(* PLC project Palletizer_Cell4.project, CODESYS CODESYS V3.5 SP19 Patch 2 *)
(* stored: creationDateTime 2026-10-30T09:14:22.5521931, modificationDateTime 2026-10-30T09:13:58.1180274 *)

(* Palletizer cell state *)
{attribute 'strict'}
TYPE E_CellState : (Idle := 0, Homing := 1, Picking := 2, Placing := 3, Faulted := 99) INT;
END_TYPE

TYPE ST_Recipe : STRUCT
  sName : STRING(40);  (* Recipe name *)
  iLayers : INT;  (* Layers per pallet *)
  iBoxesPerLayer : INT;
  lrLayerHeight : LREAL;  (* mm *)
  ltSettle : LTIME;  (* Settle time after place *)
END_STRUCT;
END_TYPE

TYPE U_StatusWord : union;
END_TYPE

INTERFACE I_Station
END_INTERFACE

FUNCTION_BLOCK ABSTRACT FB_Station IMPLEMENTS I_Station
VAR_INPUT
	bEnable : BOOL;
END_VAR
VAR_OUTPUT
	bReady : BOOL;
	nErrorId : UDINT;
END_VAR
VAR
	bFaulted : BOOL;
END_VAR

bReady := bEnable AND NOT bFaulted;

METHOD Reset : BOOL
THIS^.bFaulted := FALSE;
THIS^.nErrorId := 0;
Reset := TRUE;
END_METHOD

PROPERTY IsFaulted : BOOL
GET
IsFaulted := bFaulted;
END_GET
END_PROPERTY
END_FUNCTION_BLOCK

FUNCTION_BLOCK FB_Conveyor EXTENDS FB_Station
VAR_INPUT
	bBoxAtEnd : BOOL; // Photo-eye at discharge end
	bRunReq : BOOL;
END_VAR
VAR_OUTPUT
	bMotorOn : BOOL;
END_VAR
VAR
	tJam : TON;
	uStatus : U_StatusWord;
	fbBlink : Util.BLINK;
END_VAR

SUPER^();

// Jam: motor running but box never leaves the photo-eye
tJam(IN := bMotorOn AND bBoxAtEnd, PT := T#8S);
bFaulted S= tJam.Q;

bMotorOn := bReady AND bRunReq AND NOT bBoxAtEnd;

uStatus.wRaw.0 := bMotorOn;
uStatus.wRaw.1 := bFaulted;
uStatus.wRaw.3 := tJam.Q;

fbBlink(ENABLE := bFaulted, TIMELOW := T#500MS, TIMEHIGH := T#500MS);
END_FUNCTION_BLOCK

FUNCTION_BLOCK FB_PickAxis EXTENDS FB_Station
VAR_INPUT
	lrTargetPos : LREAL; // mm
	bMove : BOOL;
END_VAR
VAR_OUTPUT
	bInPos : BOOL;
END_VAR
VAR_IN_OUT
	Axis : AXIS_REF_SM3;
END_VAR
VAR
	fbPower : MC_Power;
	fbHome : MC_Home;
	fbMove : MC_MoveAbsolute;
END_VAR

SUPER^();
fbPower(Axis := Axis, Enable := bEnable, bRegulatorOn := bEnable, bDriveStart := bEnable);
fbHome(Axis := Axis, Execute := fbPower.Status AND NOT fbHome.Done, Position := 0);
fbMove(Axis := Axis, Execute := bMove AND fbHome.Done, Position := lrTargetPos, Velocity := 400, Acceleration := 2000, Deceleration := 2000);
bInPos := fbMove.Done;
IF fbMove.Error OR fbPower.Error THEN
	bFaulted := TRUE;
	nErrorId := fbMove.ErrorID;
END_IF
END_FUNCTION_BLOCK

{attribute 'enable_dynamic_creation'}
FUNCTION_BLOCK FB_CycleLogger
VAR_INPUT
	bLog : BOOL;
	sLine : STRING(80);
END_VAR
VAR
	hFile : FILE.CAA.HANDLE;
	fbOpen : FILE.Open;
	fbWrite : FILE.Write;
	pBuffer : POINTER TO BYTE;
	udiLen : UDINT;
	dtNow : DT;
	rtLog : R_TRIG;
END_VAR

rtLog(CLK := bLog);
IF rtLog.Q THEN
	dtNow := SysTimeRtcGet(udiLen);
	__TRY
		pBuffer := __NEW(BYTE, 128);
		udiLen := TO_UDINT(LEN(sLine));
		SysMemCpy(pBuffer, ADR(sLine), udiLen);
		fbWrite(hFile := hFile, pBuffer := pBuffer, szSize := udiLen, xExecute := TRUE);
	__CATCH
		udiLen := 0;
	__ENDTRY
	__DELETE(pBuffer);
END_IF
fbOpen(sFileName := '/data/cycles.csv', eFileMode := FILE.MODE.MAPPD, xExecute := NOT fbOpen.xDone);
hFile := fbOpen.hFile;
END_FUNCTION_BLOCK

FUNCTION_BLOCK FB_LayerCounter
  VAR_INPUT
    bBoxPlaced : BOOL;  (* Pulse when a box is released *)
    iBoxesPerLayer : INT;
    iLayers : INT;
    bReset : BOOL;
  END_VAR
  VAR_OUTPUT
    iBox : INT;
    iLayer : INT;
    bPalletFull : BOOL;
  END_VAR
  VAR
    rtBox : R_TRIG;
  END_VAR

(* Counts boxes per layer and layers per pallet *)
rtBox(CLK := bBoxPlaced);
IF bReset THEN
	iBox := 0;
	iLayer := 0;
ELSIF rtBox.Q AND NOT bPalletFull THEN
	iBox := iBox + 1;
	IF iBox >= iBoxesPerLayer THEN
		iBox := 0;
		iLayer := iLayer + 1;
	END_IF
END_IF
bPalletFull := iLayer >= iLayers;
END_FUNCTION_BLOCK

PROGRAM PLC_PRG
  VAR
    eState : E_CellState;
    fbInfeed : FB_Conveyor;
    fbAxisZ : FB_PickAxis;
    fbLog : FB_CycleLogger;
    itfStations : ARRAY[0..1] OF I_Station;
    iLayer : INT;
    iBox : INT;
    i : INT;
  END_VAR

itfStations[0] := fbInfeed;
itfStations[1] := fbAxisZ;

fbInfeed(bEnable := GVL_IO.bAutoMode, bBoxAtEnd := GVL_IO.bPE_Infeed, bRunReq := eState = E_CellState.Picking);
fbAxisZ(bEnable := GVL_IO.bAutoMode, Axis := AxisZ, lrTargetPos := GVL_Recipe.stActive.lrLayerHeight * iLayer);
GVL_IO.bConveyorMotor := fbInfeed.bMotorOn;

CASE eState OF
E_CellState.Idle:
	IF GVL_IO.bStartPB AND GVL_IO.bAutoMode THEN
		eState := E_CellState.Homing;
	END_IF
E_CellState.Homing:
	IF fbAxisZ.bReady THEN
		eState := E_CellState.Picking;
	END_IF
E_CellState.Picking:
	IF GVL_IO.bPE_Infeed THEN
		fbAxisZ.bMove := TRUE;
		eState := E_CellState.Placing;
	END_IF
E_CellState.Placing:
	IF fbAxisZ.bInPos THEN
		fbAxisZ.bMove := FALSE;
		iBox := iBox + 1;
		IF iBox >= GVL_Recipe.stActive.iBoxesPerLayer THEN
			iBox := 0;
			iLayer := iLayer + 1;
		END_IF
		fbLog(bLog := TRUE, sLine := CONCAT('box placed, layer ', INT_TO_STRING(iLayer)));
		eState := E_CellState.Picking;
	END_IF
E_CellState.Faulted:
	IF GVL_IO.bResetPB THEN
		FOR i := 0 TO 1 DO
			itfStations[i].Reset();
		END_FOR
		eState := E_CellState.Idle;
	END_IF
END_CASE

IF fbInfeed.IsFaulted OR fbAxisZ.IsFaulted THEN
	eState := E_CellState.Faulted;
END_IF
GVL_IO.bFaultLamp := eState = E_CellState.Faulted;
END_PROGRAM

PROGRAM PRG_Lamps
  VAR
    fbFlash : Util.BLINK;
  END_VAR

(* CFC diagram, written out as Structured Text *)
fbFlash(ENABLE := GVL_IO.bFaultLamp);
GVL_IO.bBeacon := fbFlash.OUT;
END_PROGRAM

PROGRAM PRG_SafetyMonitor
  VAR
    fbEStop : SF_EmergencyStop;
  END_VAR

fbEStop(Activate := TRUE, S_EStopIn := GVL_IO.bEStopChannelA, S_StartReset := FALSE, Reset := GVL_IO.bResetPB);
GVL_IO.bSafeToRun := fbEStop.S_EStopOut;
END_PROGRAM

CONFIGURATION Device
  RESOURCE Application ON PLC
    {attribute 'qualified_only'}
    VAR_GLOBAL  (* GVL_IO *)
      bStartPB AT %IX0.0 : BOOL;  (* Start pushbutton *)
      bResetPB AT %IX0.1 : BOOL;  (* Fault reset pushbutton *)
      bAutoMode AT %IX0.2 : BOOL;  (* Auto/manual selector, auto *)
      bPE_Infeed AT %IX0.3 : BOOL;  (* Infeed photo-eye *)
      bEStopChannelA AT %IX1.0 : BOOL;  (* E-stop channel A *)
      bConveyorMotor AT %QX0.0 : BOOL;  (* Infeed conveyor contactor *)
      bFaultLamp AT %QX0.1 : BOOL;
      bBeacon AT %QX0.2 : BOOL;
      bSafeToRun : BOOL;
    END_VAR
    {attribute 'qualified_only'}
    VAR_GLOBAL PERSISTENT  (* GVL_Recipe *)
      stActive : ST_Recipe;
      udiPalletsDone : UDINT;
    END_VAR
    TASK EtherCAT_Task(INTERVAL := T#2ms, PRIORITY := 0);
    TASK MainTask(INTERVAL := T#10ms, PRIORITY := 1);
    TASK LogTask(INTERVAL := T#200ms, PRIORITY := 20);
    PROGRAM PRG_Motion WITH EtherCAT_Task : PRG_Motion;
    PROGRAM PLC_PRG WITH MainTask : PLC_PRG;
    PROGRAM PRG_Lamps WITH MainTask : PRG_Lamps;
    PROGRAM PRG_SafetyMonitor WITH LogTask : PRG_SafetyMonitor;
  END_RESOURCE
END_CONFIGURATION
